INTERFACE I_Fuse

PROPERTY inError : BOOL
GET
END_GET
END_PROPERTY

END_INTERFACE

(* stored: Version 1.1.0.1, ProductVersion 3.1.4024.12
   Itf I_Fuse: Id {258316fe-bb84-4bf0-b022-b1181887a622}
   Property inError: Id {8131d4f1-99f9-4d71-9dbf-63381a3ca8f5}
   Get Get: Id {e3e0986c-4202-473b-9b83-803d3a832a09} *)
